FUNCTION_BLOCK RASPBERRY_PI_CONTROL_ROBOT
  {SET_ATTRIBUTE(OpcUa, POINT.STARTPOINT)}
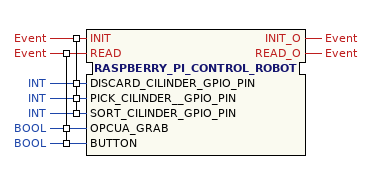
  EVENT_INPUT
    INIT WITH DISCARD_CILINDER_GPIO_PIN, PICK_CILINDER__GPIO_PIN, SORT_CILINDER_GPIO_PIN;
    READ WITH OPCUA_GRAB, BUTTON;
  END_EVENT
  EVENT_OUTPUT
    INIT_O;
    READ_O;
  END_EVENT
  VAR_INPUT
    DISCARD_CILINDER_GPIO_PIN : INT; {SET_ATTRIBUTE(OpcUa, Constant.RUN)}
    PICK_CILINDER__GPIO_PIN : INT; {SET_ATTRIBUTE(OpcUa, Constant.RUN)}
    SORT_CILINDER_GPIO_PIN : INT; {SET_ATTRIBUTE(OpcUa, Constant.RUN)}
    OPCUA_GRAB : BOOL; {SET_ATTRIBUTE(OpcUa, Variable.RUN)}
    BUTTON : BOOL; {SET_ATTRIBUTE(OpcUa, Variable.RUN)}
  END_VAR
END_FUNCTION_BLOCK
